Fanuc KAREL source: KT00842.KL

PROGRAM KT00842
%NOLOCKGROUP
VAR
  S1: STRING[80]
  S2: STRING[80]
  OUT: INTEGER
BEGIN
  S1 = 'A'
  S2 = 'B'
  S1 = 'A'
  S2 = 'B'
  OUT = SQRT(S1)
END KT00842
